Fanuc KAREL source: KD00032.KL

PROGRAM KD00032
%NOLOCKGROUP
VAR
  I: INTEGER
  J: INTEGER
  B: BOOLEAN
  R: REAL
  S: STRING[80]
BEGIN
  CONDITION[1]:
  WHEN ERROR[11038] DO
    I = 1
  ENDCONDITION
END KD00032
